FUNCTION_BLOCK UCT_Equipamento (* Equipamento de uma UCT (so IHM) - HidrycoLib *)
  (* Standard: 61499-2 *)
  (* Version 1.5, 03/11/2026, Hidryco, Hidryco, 1.5: IThis com nomes do Citect (CMD_MANUAL, STP_VELOCIDADE, CMD_INTERMITENTE, HABILITA_REVERSAO, STS_HORIMETRO_HOR); interface do CAT igual. 1.4: motor da rosca inclinada virado para a calha, A/M centralizado na caixa. 1.3: simbolos no padrao do Motor_Generico (graficos da HidrycoLib com Animacao e cores HidrycoColors, falha de comunicacao, A/M, nome), formas sobrepostas na ordem certa, area do simbolo (SymbolSize). 1.2: simbolos graficos por tipo de equipamento (sPeneira, sBomba, sValvula, sRosca, sRoscaInclinada, sCompressor, sRaspador) para o desenho do skid. 1.0: simbolo e faceplate de um equipamento da UCT Fast (peneira, bombas e valvulas de higienizacao, compressor, raspador, roscas). Recebe o estado lido da UCT pelo CAT UCT_PreTratamento e devolve os comandos da IHM (liga manual, velocidade, intermitente, reversao), um evento por comando. Nomes do IThis iguais aos dos CATs antigos da biblioteca. *)
  PACKAGE Hidryco.HidrycoLib;
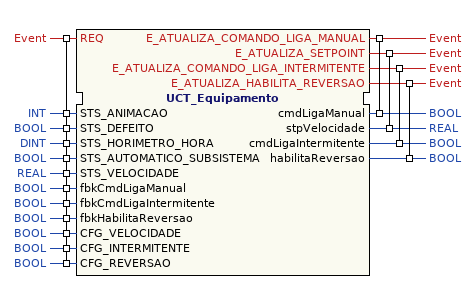
  EVENT_INPUT
    REQ WITH STS_ANIMACAO, STS_DEFEITO, STS_HORIMETRO_HORA, STS_AUTOMATICO_SUBSISTEMA, STS_VELOCIDADE, fbkCmdLigaManual, fbkCmdLigaIntermitente, fbkHabilitaReversao, CFG_VELOCIDADE, CFG_INTERMITENTE, CFG_REVERSAO; (* Estado da UCT *)
  END_EVENT
  EVENT_OUTPUT
    E_ATUALIZA_COMANDO_LIGA_MANUAL WITH cmdLigaManual; (* IHM: liga (TRUE) / desliga (FALSE) em manual *)
    E_ATUALIZA_SETPOINT WITH stpVelocidade; (* IHM: velocidade (%) *)
    E_ATUALIZA_COMANDO_LIGA_INTERMITENTE WITH cmdLigaIntermitente; (* IHM: liga (TRUE) / desliga (FALSE) o intermitente *)
    E_ATUALIZA_HABILITA_REVERSAO WITH habilitaReversao; (* IHM: habilita (TRUE) / desabilita (FALSE) a reversao *)
  END_EVENT
  VAR_INPUT
    STS_ANIMACAO : INT; (* Estado do equipamento na UCT: 0 desligado, 1 ligado, 2 falha, 3 manutencao, 4 sem comunicacao *)
    STS_DEFEITO : BOOL; (* Defeito do equipamento (palavra 40081 da UCT) *)
    STS_HORIMETRO_HORA : DINT; (* Horimetro do equipamento (h, lido da UCT) *)
    STS_AUTOMATICO_SUBSISTEMA : BOOL; (* Subsistema do equipamento em automatico (comandos manuais bloqueados) *)
    STS_VELOCIDADE : REAL; (* Velocidade ajustada na UCT (%) *)
    fbkCmdLigaManual : BOOL; (* Comando liga em vigor na UCT *)
    fbkCmdLigaIntermitente : BOOL; (* Modo intermitente em vigor na UCT *)
    fbkHabilitaReversao : BOOL; (* Reversao habilitada na UCT *)
    CFG_VELOCIDADE : BOOL; (* TRUE = equipamento com ajuste de velocidade *)
    CFG_INTERMITENTE : BOOL; (* TRUE = equipamento com modo intermitente *)
    CFG_REVERSAO : BOOL; (* TRUE = equipamento com reversao *)
  END_VAR
  VAR_OUTPUT
    cmdLigaManual : BOOL; (* IHM: liga (TRUE) / desliga (FALSE) em manual *)
    stpVelocidade : REAL; (* IHM: velocidade (%) *)
    cmdLigaIntermitente : BOOL; (* IHM: liga (TRUE) / desliga (FALSE) o intermitente *)
    habilitaReversao : BOOL; (* IHM: habilita (TRUE) / desabilita (FALSE) a reversao *)
  END_VAR
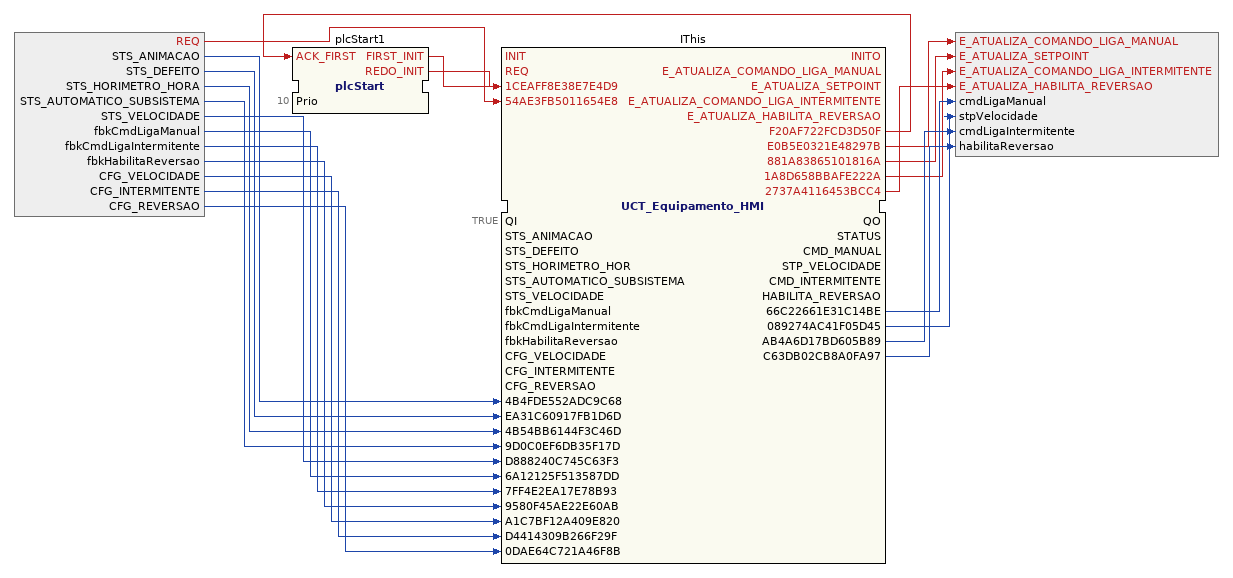
  FBS
    IThis : UCT_Equipamento_HMI(QI := TRUE);
    plcStart1 : plcStart(Prio := 10);
  END_FBS
  EVENT_CONNECTIONS
    plcStart1.FIRST_INIT TO IThis.1CEAFF8E38E7E4D9;
    plcStart1.REDO_INIT TO IThis.1CEAFF8E38E7E4D9;
    IThis.F20AF722FCD3D50F TO plcStart1.ACK_FIRST;
    REQ TO IThis.54AE3FB5011654E8;
    IThis.E0B5E0321E48297B TO E_ATUALIZA_COMANDO_LIGA_MANUAL;
    IThis.881A83865101816A TO E_ATUALIZA_SETPOINT;
    IThis.1A8D658BBAFE222A TO E_ATUALIZA_COMANDO_LIGA_INTERMITENTE;
    IThis.2737A4116453BCC4 TO E_ATUALIZA_HABILITA_REVERSAO;
  END_CONNECTIONS
  DATA_CONNECTIONS
    STS_ANIMACAO TO IThis.4B4FDE552ADC9C68;
    STS_DEFEITO TO IThis.EA31C60917FB1D6D;
    STS_HORIMETRO_HORA TO IThis.4B54BB6144F3C46D;
    STS_AUTOMATICO_SUBSISTEMA TO IThis.9D0C0EF6DB35F17D;
    STS_VELOCIDADE TO IThis.D888240C745C63F3;
    fbkCmdLigaManual TO IThis.6A12125F513587DD;
    fbkCmdLigaIntermitente TO IThis.7FF4E2EA17E78B93;
    fbkHabilitaReversao TO IThis.9580F45AE22E60AB;
    CFG_VELOCIDADE TO IThis.A1C7BF12A409E820;
    CFG_INTERMITENTE TO IThis.D4414309B266F29F;
    CFG_REVERSAO TO IThis.0DAE64C721A46F8B;
    IThis.66C22661E31C14BE TO cmdLigaManual;
    IThis.089274AC41F05D45 TO stpVelocidade;
    IThis.AB4A6D17BD605B89 TO cmdLigaIntermitente;
    IThis.C63DB02CB8A0FA97 TO habilitaReversao;
  END_CONNECTIONS
END_FUNCTION_BLOCK
